(* IEC 61131-3 sources: plcassist-cli/packages/volt-lsp-iec/test-corpus/bakon-nano/Device/Plc Logic/Application/Library Manager/L_IE1P_ApplicationErrorsTypes, 11 files *)

(* ---- GVL.gvl ---- *)
VAR_GLOBAL
END_VAR

(* ---- L_IE1P_IERRORHANDLER.itf ---- *)
INTERFACE L_IE1P_IERRORHANDLER
END_INTERFACE

METHOD ITFCHECKERRORRESETOCCURED : BOOL
VAR_IN_OUT
	RESETTIME : SYSTIME;
END_VAR
END_METHOD

METHOD ITFCLEARERROR : DWORD
VAR_INPUT
	ESEVERITY : L_IE1P_SeverityLevel;
	WERRORID : WORD;
	WCOMPID : WORD;
	DWINSTANCEID : DWORD := 0;
END_VAR
END_METHOD

METHOD ITFCLEARREACTION
VAR_INPUT
	EREACTION : L_IE1P_Reaction;
	DICLEARCOUNT : DINT;
	DWINSTANCEID : DWORD;
END_VAR
END_METHOD

METHOD ITFGETACTUALERRORCODE : DWORD
VAR_OUTPUT
	ESEVERITY : WORD;
END_VAR
END_METHOD

METHOD ITFREGISTERERRORINSTANCE : DWORD
END_METHOD

METHOD ITFRESETACTIVE : BOOL
END_METHOD

METHOD ITFRESETERROR : DWORD
VAR_INPUT
	ERRORHANDLE : RTS_IEC_HANDLE := 0;
END_VAR
END_METHOD

METHOD ITFRESETERRORREACTION
VAR_INPUT
	DWINSTANCEID : DWORD := 0;
END_VAR
END_METHOD

METHOD ITFSETERROR : DWORD
VAR_INPUT
	ESEVERITY : L_IE1P_SeverityLevel;
	WERRORID : WORD;
	WCOMPID : WORD;
	DWINSTANCEID : DWORD := 0;
	EREACTION : L_IE1P_Reaction;
END_VAR
END_METHOD

(* ---- GETBOOLEANPROPERTY.fun ---- *)
FUNCTION GETBOOLEANPROPERTY : BOOL
VAR_INPUT
	STKEY : WSTRING;
END_VAR
END_FUNCTION

(* ---- GETCOMPANY.fun ---- *)
FUNCTION GETCOMPANY : WSTRING
END_FUNCTION

(* ---- GETNUMBERPROPERTY.fun ---- *)
FUNCTION GETNUMBERPROPERTY : DINT
VAR_INPUT
	STKEY : WSTRING;
END_VAR
END_FUNCTION

(* ---- GETTEXTPROPERTY.fun ---- *)
FUNCTION GETTEXTPROPERTY : WSTRING
VAR_INPUT
	STKEY : WSTRING;
END_VAR
END_FUNCTION

(* ---- GETTEXTPROPERTY2.fun ---- *)
FUNCTION GETTEXTPROPERTY2 : POINTER TO WSTRING
VAR_INPUT
	STKEY : WSTRING;
END_VAR
END_FUNCTION

(* ---- GETTITLE.fun ---- *)
FUNCTION GETTITLE : WSTRING
END_FUNCTION

(* ---- GETVERSION.fun ---- *)
FUNCTION GETVERSION : VERSION
END_FUNCTION

(* ---- GETVERSIONPROPERTY.fun ---- *)
FUNCTION GETVERSIONPROPERTY : VERSION
VAR_INPUT
	STKEY : WSTRING;
END_VAR
END_FUNCTION

(* ---- LENZEERRMGR_11264.fb ---- *)
FUNCTION_BLOCK LENZEERRMGR_11264
VAR
	M_TEXTLISTFILE : STRING(255);
	_STNAMESPACE : STRING;
END_VAR
END_FUNCTION_BLOCK
